(* IEC 61131-3 sources: llm-plc-st-eval/data/definitivo/gpt-4o-2024-08-06/I1/zero_shot, 3 files *)

(* ---- ejec_1.st ---- *)
```pascal
FUNCTION_BLOCK FB_Semaforo
VAR_INPUT
    habilitado : BOOL; // Entrada para habilitar o deshabilitar el semáforo
END_VAR_INPUT

VAR_OUTPUT
    luzV : BOOL; // Salida para la luz verde
    luzA : BOOL; // Salida para la luz amarilla
    luzR : BOOL; // Salida para la luz roja
END_VAR_OUTPUT

VAR
    estado : INT; // Estado actual del semáforo
    temporizador : TON; // Temporizador para controlar los tiempos de las luces
    parpadeo : BOOL; // Estado del parpadeo amarillo
END_VAR

// Inicialización del bloque de función
IF NOT habilitado THEN
    // Si no está habilitado, activar parpadeo amarillo
    luzV := FALSE;
    luzR := FALSE;
    temporizador(IN := TRUE, PT := T#1S);
    parpadeo := temporizador.Q;
    luzA := parpadeo;
ELSE
    // Si está habilitado, seguir la secuencia normal del semáforo
    temporizador(IN := TRUE);
    CASE estado OF
        0: // Luz verde
            luzV := TRUE;
            luzA := FALSE;
            luzR := FALSE;
            temporizador(PT := T#20S);
            IF temporizador.Q THEN
                estado := 1;
                temporizador(IN := FALSE);
            END_IF;
        1: // Luz amarilla
            luzV := FALSE;
            luzA := TRUE;
            luzR := FALSE;
            temporizador(PT := T#4S);
            IF temporizador.Q THEN
                estado := 2;
                temporizador(IN := FALSE);
            END_IF;
        2: // Luz roja
            luzV := FALSE;
            luzA := FALSE;
            luzR := TRUE;
            temporizador(PT := T#15S);
            IF temporizador.Q THEN
                estado := 0;
                temporizador(IN := FALSE);
            END_IF;
    ELSE
        // Reiniciar al estado inicial si el estado es desconocido
        estado := 0;
    END_CASE;
END_IF;
END_FUNCTION_BLOCK
```

Este código implementa un semáforo vehicular cíclico en un bloque de función `FB_Semaforo` usando Structured Text (ST) conforme al estándar IEC 61131-3. El semáforo sigue una secuencia de luces verde, amarilla y roja cuando está habilitado, y cambia a un parpadeo amarillo cuando está deshabilitado.

(* ---- ejec_2.st ---- *)
```pascal
FUNCTION_BLOCK FB_Semaforo
VAR
    // Variables de entrada
    habilitado : BOOL; // Entrada para habilitar o deshabilitar el semáforo

    // Variables de salida
    luzV : BOOL; // Luz verde
    luzA : BOOL; // Luz amarilla
    luzR : BOOL; // Luz roja

    // Variables internas
    estado : INT := 0; // Estado del semáforo
    temporizador : TON; // Temporizador para controlar los tiempos de las luces
    tiempoParpadeo : TON; // Temporizador para el parpadeo del amarillo
END_VAR

// Inicialización del temporizador
temporizador(IN := FALSE, PT := T#0S);
tiempoParpadeo(IN := FALSE, PT := T#0S);

// Lógica del semáforo
IF habilitado THEN
    // Secuencia cíclica del semáforo
    CASE estado OF
        0: // Luz verde
            luzV := TRUE;
            luzA := FALSE;
            luzR := FALSE;
            temporizador(IN := TRUE, PT := T#20S);
            IF temporizador.Q THEN
                temporizador(IN := FALSE);
                estado := 1;
            END_IF;
        1: // Luz amarilla
            luzV := FALSE;
            luzA := TRUE;
            luzR := FALSE;
            temporizador(IN := TRUE, PT := T#4S);
            IF temporizador.Q THEN
                temporizador(IN := FALSE);
                estado := 2;
            END_IF;
        2: // Luz roja
            luzV := FALSE;
            luzA := FALSE;
            luzR := TRUE;
            temporizador(IN := TRUE, PT := T#15S);
            IF temporizador.Q THEN
                temporizador(IN := FALSE);
                estado := 0;
            END_IF;
    END_CASE;
ELSE
    // Modo amarillo intermitente
    luzV := FALSE;
    luzR := FALSE;
    tiempoParpadeo(IN := TRUE, PT := T#1S);
    IF tiempoParpadeo.Q THEN
        luzA := NOT luzA; // Alterna el estado de la luz amarilla
        tiempoParpadeo(IN := FALSE);
    END_IF;
    estado := 0; // Reinicia el estado para comenzar en verde cuando se habilite
END_IF;
END_FUNCTION_BLOCK
```

(* ---- ejec_3.st ---- *)
```pascal
FUNCTION_BLOCK FB_Semaforo
VAR_INPUT
    habilitado : BOOL; // Entrada para habilitar o deshabilitar el semáforo
END_VAR_INPUT

VAR_OUTPUT
    luzV : BOOL; // Salida para la luz verde
    luzA : BOOL; // Salida para la luz amarilla
    luzR : BOOL; // Salida para la luz roja
END_VAR_OUTPUT

VAR
    estado : INT := 0; // Estado del semáforo
    temporizador : TON; // Temporizador para manejar los tiempos
    parpadeo : BOOL := FALSE; // Estado del parpadeo amarillo
END_VAR

// Inicialización del temporizador
temporizador(IN := FALSE, PT := T#0S);

IF habilitado THEN
    // Secuencia cíclica del semáforo
    CASE estado OF
        0: // Luz verde
            luzV := TRUE;
            luzA := FALSE;
            luzR := FALSE;
            temporizador(IN := TRUE, PT := T#20S);
            IF temporizador.Q THEN
                estado := 1;
                temporizador(IN := FALSE);
            END_IF;
        1: // Luz amarilla
            luzV := FALSE;
            luzA := TRUE;
            luzR := FALSE;
            temporizador(IN := TRUE, PT := T#4S);
            IF temporizador.Q THEN
                estado := 2;
                temporizador(IN := FALSE);
            END_IF;
        2: // Luz roja
            luzV := FALSE;
            luzA := FALSE;
            luzR := TRUE;
            temporizador(IN := TRUE, PT := T#15S);
            IF temporizador.Q THEN
                estado := 0;
                temporizador(IN := FALSE);
            END_IF;
    END_CASE;
ELSE
    // Modo amarillo intermitente
    luzV := FALSE;
    luzR := FALSE;
    temporizador(IN := TRUE, PT := T#1S);
    IF temporizador.Q THEN
        parpadeo := NOT parpadeo;
        temporizador(IN := FALSE);
    END_IF;
    luzA := parpadeo;
    estado := 0; // Reiniciar secuencia al habilitar
END_IF;
END_FUNCTION_BLOCK
```

Este código implementa un semáforo vehicular cíclico en un bloque de función llamado `FB_Semaforo`. Utiliza un temporizador para controlar la duración de cada luz y cambia de estado según el tiempo transcurrido. Cuando la entrada `habilitado` está desactivada, el semáforo entra en un modo de parpadeo amarillo. Al reactivarse, la secuencia comienza nuevamente con la luz verde.
